FUNCTION_BLOCK ARM_Control (* Basic Function Block Type *)
  (* Standard: 61499-2 *)
  (* Version 0.0, 10/20/2026, lizar, Schneider Electric, Template *)
  PACKAGE Main;
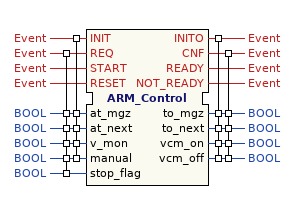
  EVENT_INPUT
    INIT WITH at_mgz, at_next, v_mon, manual; (* Initialization Request *)
    REQ WITH at_mgz, at_next, v_mon, manual, stop_flag; (* Normal Execution Request *)
    START;
    RESET;
  END_EVENT
  EVENT_OUTPUT
    INITO WITH to_mgz, to_next, vcm_on, vcm_off; (* Initialization Confirm *)
    CNF WITH to_mgz, to_next, vcm_on, vcm_off; (* Execution Confirmation *)
    READY;
    NOT_READY;
  END_EVENT
  VAR_INPUT
    at_mgz : BOOL; (* Input event qualifier *)
    at_next : BOOL;
    v_mon : BOOL;
    manual : BOOL;
    stop_flag : BOOL;
  END_VAR
  VAR_OUTPUT
    to_mgz : BOOL; (* Output event qualifier *)
    to_next : BOOL;
    vcm_on : BOOL;
    vcm_off : BOOL;
  END_VAR
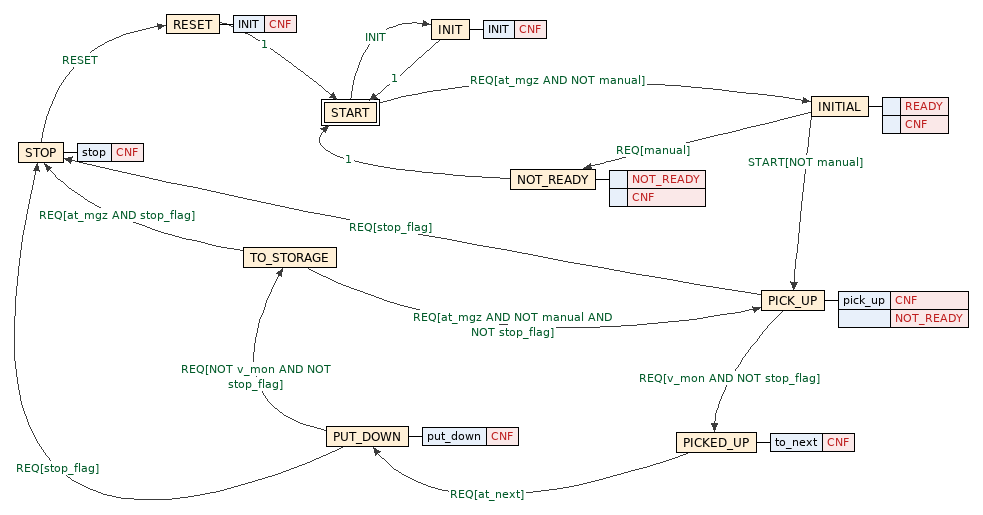
  EC_STATES
    START; (* Initial State *)
    INIT : INIT -> CNF; (* Initialization *)
    INITIAL : -> READY, -> CNF;
    PICK_UP : pick_up -> CNF, -> NOT_READY;
    PUT_DOWN : put_down -> CNF;
    PICKED_UP : to_next -> CNF;
    TO_STORAGE;
    NOT_READY : -> NOT_READY, -> CNF;
    STOP : stop -> CNF;
    RESET : INIT -> CNF;
  END_STATES
  EC_TRANSITIONS
    START TO INIT := INIT;
    INIT TO START := 1;
    START TO INITIAL := REQ[at_mgz AND NOT manual];
    INITIAL TO PICK_UP := START[NOT manual];
    PICKED_UP TO PUT_DOWN := REQ[at_next];
    TO_STORAGE TO PICK_UP := REQ[at_mgz AND NOT manual AND NOT stop_flag];
    PICK_UP TO PICKED_UP := REQ[v_mon AND NOT stop_flag];
    PUT_DOWN TO TO_STORAGE := REQ[NOT v_mon AND NOT stop_flag];
    INITIAL TO NOT_READY := REQ[manual];
    NOT_READY TO START := 1;
    PUT_DOWN TO STOP := REQ[stop_flag];
    TO_STORAGE TO STOP := REQ[at_mgz AND stop_flag];
    RESET TO START := 1;
    STOP TO RESET := RESET;
    PICK_UP TO STOP := REQ[stop_flag];
  END_TRANSITIONS
  ALGORITHM INIT IN ST: (* Initialization algorithm *)
;
to_mgz:=TRUE;
to_next:=FALSE;
vcm_off:=TRUE;
vcm_on:=FALSE;
  END_ALGORITHM
  ALGORITHM pick_up IN ST:
;
vcm_on:=TRUE;
vcm_off:=FALSE;
  END_ALGORITHM
  ALGORITHM put_down IN ST:
;
vcm_on:=FALSE;
vcm_off:=TRUE;
to_mgz:=TRUE;
to_next:= FALSE;
  END_ALGORITHM
  ALGORITHM to_next IN ST:
;
to_mgz:=FALSE;
to_next:=TRUE;
  END_ALGORITHM
  ALGORITHM stop IN ST:
;
to_mgz:=FALSE;
to_next:=FALSE;
vcm_on:=FALSE;
vcm_off:=TRUE;
  END_ALGORITHM
END_FUNCTION_BLOCK
